// TIA Portal V21 export
// export: Created 2026-10-24T16:33:10.0564923Z, ExportSetting WithDefaults, DisplayName Totally Integrated Automation Portal, DisplayVersion V21 Update 1, DisplayName SINAMICS Startdrive Advanced, DisplayVersion V21 HF2, DisplayName SINAMICS Startdrive G110M, G120, G120C, G120D, G120P, G115D, DisplayVersion V21 HF2, DisplayName SINAMICS Startdrive G130, G150, S120, S150, G200, G220, S200, S210, S220, Innomotics MVD, DisplayVersion V21 HF2, DisplayName STEP 7 Professional, DisplayVersion V21 Update 1, DisplayName STEP 7 Safety, DisplayVersion V21, DisplayName Tech WebApplication, DisplayVersion V21, DisplayName WinCC Basic/Comfort/Advanced, DisplayVersion V21 Update 1, DisplayName WinCC Unified, DisplayVersion V21 Update 1
FUNCTION_BLOCK "FB_V4_Tally"   // FB37, SCL
{ S7_Optimized_Access := 'TRUE' }
VERSION : 0.1
// stored: AutoNumber true, IsIECCheckEnabled false, IsRetainMemResEnabled false, MemoryReserve 100, SetENOAutomatically false, UDAEnableTagReadback false
   VAR_INPUT
      Execute : Bool;   // Count on every call while true
   END_VAR
   VAR_OUTPUT
      Count : Int;   // Calls counted
   END_VAR
   VAR
      Tally { S7_SetPoint := 'True'} : "UDT_V4_Counter";   // Internal tally
   END_VAR
BEGIN

       IF #Execute THEN
           "FC_V4_Advance"(Tally := #Tally);
       END_IF;
       #Count := #Tally.Count;
END_FUNCTION_BLOCK
